(* IEC 61131-3 sources: nautilus/internal/project/testdata/libdir/lib, 1 file *)

(* ---- blocks.st ---- *)
FUNCTION_BLOCK HiAlarm
VAR_INPUT
    PV : REAL;
    Limit : REAL;
END_VAR
VAR_OUTPUT
    Alm : BOOL;
END_VAR
Alm := PV > Limit;
END_FUNCTION_BLOCK
